{attribute 'qualified_only'}
{attribute 'strict'}
TYPE E_UmTutorialCmd :
(
	NoCmd
);
END_TYPE

(* stored: Version 1.1.0.1, ProductVersion 3.1.4024.12
   DUT E_UmTutorialCmd: Id {0cd378ee-6ee8-4531-acd8-ff5b30a7272b} *)
